// TIA Portal project "072_motion_tcpu" (V21)

(* hardware
DEVICE "PLC_T"  S7-1500 station
   slot 0: "Rail_0"  Rack  6ES7 590-1***0-0AA0
   slot 1: "PLC_T"  CPU 1515T-2 PN  6ES7 515-2TN03-0AB0  V3.1
      slot 3: "CPU display_1"  6ES7591-1BA00-0AA0
      slot 32768: "PROFINET interface_1"  X1
         slot 32769: "Port_1"  X1 P1
         slot 32770: "Port_2"  X1 P2
      slot 33024: "PROFINET interface_2"  X2
         slot 33025: "Port_1"  X2 P1
      slot 34817: "Virtual CP interface port_1"  Virtual CP interface port  Virtual CP interface port
   slot 2: "TM_Timer_1"  TM Timer DIDQ 16x24V  6ES7 552-1AA00-0AB0  V1.0
      slot 1: "TM_Timer_1"  TM Timer DIDQ 16x24V
*)

// ===== PLC "PLC_T"  CPU 1515T-2 PN =====

VAR_GLOBAL   // PLC tag table "Default tag table"
   "MeasuringInput_1_Interface_Address" AT %I0.0 : Bool;
END_VAR

DATA_BLOCK "DB_Enc"   // DB15
{ S7_Optimized_Access := 'FALSE' }
VERSION : 0.1
   VAR
      tel : PD_TEL81;
   END_VAR
BEGIN
END_DATA_BLOCK

DATA_BLOCK "mTO_PositioningAxis"   // DB1, Motion_DB
{ S7_Optimized_Access := 'TRUE' }
AUTHOR : SIMATIC
FAMILY : MC_1500
VERSION : 8.0
// stored: InstanceOfName TO_PositioningAxis
"TO_PositioningAxis"
BEGIN
END_DATA_BLOCK

DATA_BLOCK "mTO_SynchronousAxis"   // DB2, Motion_DB
{ S7_Optimized_Access := 'TRUE' }
AUTHOR : SIMATIC
FAMILY : MC_1500
VERSION : 8.0
// stored: InstanceOfName TO_SynchronousAxis
"TO_SynchronousAxis"
BEGIN
END_DATA_BLOCK

DATA_BLOCK "mTO_Cam"   // DB3, Motion_DB
{ S7_Optimized_Access := 'TRUE' }
AUTHOR : SIMATIC
FAMILY : MC_1500
VERSION : 8.0
// stored: InstanceOfName TO_Cam
"TO_Cam"
BEGIN
END_DATA_BLOCK

DATA_BLOCK "mTO_Cam_10k"   // DB4, Motion_DB
{ S7_Optimized_Access := 'TRUE' }
AUTHOR : SIMATIC
FAMILY : MC_1500
VERSION : 8.0
// stored: InstanceOfName TO_Cam_10k
"TO_Cam_10k"
BEGIN
END_DATA_BLOCK

DATA_BLOCK "mTO_LeadingAxisProxy"   // DB5, Motion_DB
{ S7_Optimized_Access := 'TRUE' }
AUTHOR : SIMATIC
FAMILY : MC_1500
VERSION : 8.0
// stored: InstanceOfName TO_LeadingAxisProxy
"TO_LeadingAxisProxy"
BEGIN
END_DATA_BLOCK

DATA_BLOCK "mTO_Kinematics"   // DB6, Motion_DB
{ S7_Optimized_Access := 'TRUE' }
AUTHOR : SIMATIC
FAMILY : MC_1500
VERSION : 8.0
// stored: InstanceOfName TO_Kinematics
"TO_Kinematics"
BEGIN
END_DATA_BLOCK

DATA_BLOCK "mTO_SpeedAxis"   // DB7, Motion_DB
{ S7_Optimized_Access := 'TRUE' }
AUTHOR : SIMATIC
FAMILY : MC_1500
VERSION : 8.0
// stored: InstanceOfName TO_SpeedAxis
"TO_SpeedAxis"
BEGIN
END_DATA_BLOCK

DATA_BLOCK "mTO_ExternalEncoder"   // DB8, Motion_DB
{ S7_Optimized_Access := 'TRUE' }
AUTHOR : SIMATIC
FAMILY : MC_1500
VERSION : 8.0
// stored: InstanceOfName TO_ExternalEncoder
"TO_ExternalEncoder"
BEGIN
END_DATA_BLOCK

DATA_BLOCK "mTO_Interpreter"   // DB9, Motion_DB
{ S7_Optimized_Access := 'TRUE' }
AUTHOR : SIMATIC
FAMILY : MC_1500
VERSION : 8.0
// stored: InstanceOfName TO_Interpreter
"TO_Interpreter"
BEGIN
END_DATA_BLOCK

DATA_BLOCK "mTO_InterpreterMapping"   // DB10, Motion_DB
{ S7_Optimized_Access := 'TRUE' }
AUTHOR : SIMATIC
FAMILY : MC_1500
VERSION : 8.0
// stored: InstanceOfName TO_InterpreterMapping
"TO_InterpreterMapping"
BEGIN
END_DATA_BLOCK

DATA_BLOCK "mTO_InterpreterProgram"   // DB11, Motion_DB
{ S7_Optimized_Access := 'TRUE' }
AUTHOR : SIMATIC
FAMILY : MC_1500
VERSION : 8.0
// stored: InstanceOfName TO_InterpreterProgram
"TO_InterpreterProgram"
BEGIN
END_DATA_BLOCK

DATA_BLOCK "OutputCam_1"   // DB12, Motion_DB
{ S7_Optimized_Access := 'TRUE' }
AUTHOR : SIMATIC
FAMILY : MC_1500
VERSION : 8.0
// stored: InstanceOfName TO_OutputCam
"TO_OutputCam"
BEGIN
END_DATA_BLOCK

DATA_BLOCK "CamTrack_1"   // DB13, Motion_DB
{ S7_Optimized_Access := 'TRUE' }
AUTHOR : SIMATIC
FAMILY : MC_1500
VERSION : 8.0
// stored: InstanceOfName TO_CamTrack
"TO_CamTrack"
BEGIN
END_DATA_BLOCK

DATA_BLOCK "MeasuringInput_1"   // DB14, Motion_DB
{ S7_Optimized_Access := 'TRUE' }
AUTHOR : SIMATIC
FAMILY : MC_1500
VERSION : 8.0
// stored: InstanceOfName TO_MeasuringInput
"TO_MeasuringInput"
BEGIN
END_DATA_BLOCK

ORGANIZATION_BLOCK "Main"   // OB1, LAD, ProgramCycle
TITLE = "Main Program Sweep (Cycle)"
{ S7_Optimized_Access := 'TRUE' }
VERSION : 0.1
   VAR_INPUT
      Initial_Call : Bool;   // Initial call of this OB
      Remanence : Bool;   // =True, if remanent data are available
   END_VAR
BEGIN
END_ORGANIZATION_BLOCK